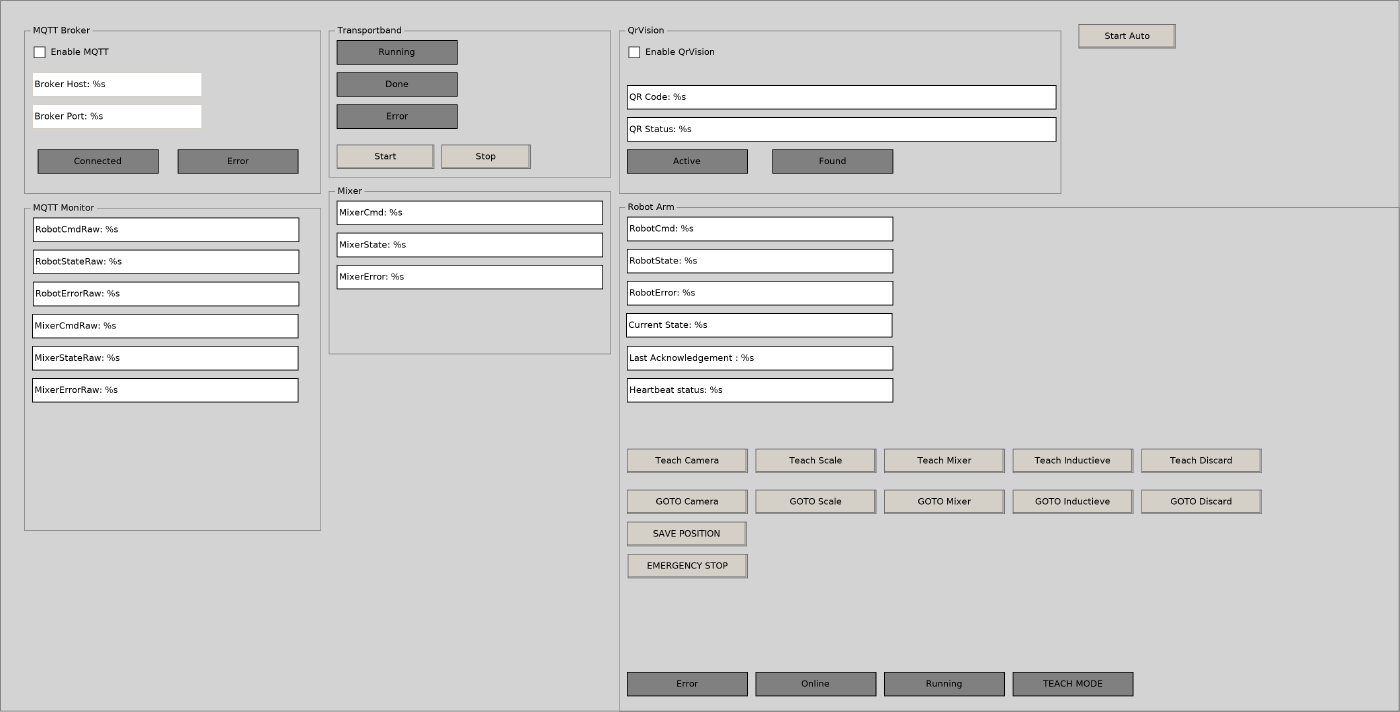
VISUALIZATION PannenkoekenDashboard  // 1742x887
    GroupBox (30,30 369x211), "MQTT Broker"
        Checkbox (10,20 150x30), "Enable MQTT", variable: GVL_MQTT.bEnableMqtt
        Rectangle (191,156 150x30), "Error"
        Rectangle (17,156 150x30), "Connected", colour toggle: GVL_MQTT.bMqttConnected
        Textfield (10,60 211x30), "Broker Host: %s", text variable: GVL_MQTT.sMqttBroker
        Textfield (10,100 211x30), "Broker Port: %s", text variable: GVL_MQTT.nMqttPort
    GroupBox (30,251 369x410), "MQTT Monitor"
        Rectangle (10,140 331x30), "MixerCmdRaw: %s", text variable: GVL_MQTT.sMixerCmdRaw
        Rectangle (10,180 331x30), "MixerStateRaw: %s", text variable: GVL_MQTT.sMixerStateRaw
        Rectangle (10,220 331x30), "MixerErrorRaw: %s", text variable: GVL_MQTT.sMixerErrorRaw
        Rectangle (11,20 331x30), "RobotCmdRaw: %s", text variable: GVL_MQTT.sRobotCmdRaw
        Rectangle (11,60 331x30), "RobotStateRaw: %s", text variable: GVL_MQTT.sRobotStateRaw
        Rectangle (11,100 331x30), "RobotErrorRaw: %s", text variable: GVL_MQTT.sRobotErrorRaw
    GroupBox (770,250 972x637), "Robot Arm"
        Rectangle (10,20 331x30), "RobotCmd: %s", text variable: GVL_MQTT.sRobotCmdDisplay
        Rectangle (10,60 331x30), "RobotState: %s", text variable: GVL_MQTT.sRobotStateDisplay
        Rectangle (10,100 331x30), "RobotError: %s", text variable: GVL_MQTT.sRobotErrorDisplay
        Rectangle (10,587 150x30), "Error", colour toggle: GVL_MQTT.bRobotArmAlarm
        Rectangle (170,587 150x30), "Online", colour toggle: GVL_MQTT.bRobotArmOnline
        Rectangle (330,587 150x30), "Running", colour toggle: GVL_MQTT.bRobotArmBusy
        Rectangle (10,221 331x30), "Heartbeat status: %s", text variable: GVL_MQTT.sRobotHeartbeatDisplay
        Rectangle (9,140 331x30), "Current State: %s", text variable: GVL_MQTT.sRobotArmDisplay
        Button (10,309 150x30), "Teach Camera"
            OnMouseClick: execute { GVL_MQTT.sRobotTargetPose := 'camera'; GVL_MQTT.bVisuRobotTeach  := TRUE; }
        Button (170,309 150x30), "Teach Scale"
            OnMouseClick: execute { GVL_MQTT.sRobotTargetPose := 'scale'; GVL_MQTT.bVisuRobotTeach  := TRUE; }
        Button (330,309 150x30), "Teach Mixer"
            OnMouseClick: execute { GVL_MQTT.sRobotTargetPose := 'mixer'; GVL_MQTT.bVisuRobotTeach  := TRUE; }
        Button (490,309 150x30), "Teach Inductieve"
            OnMouseClick: execute { GVL_MQTT.sRobotTargetPose := 'inductive'; GVL_MQTT.bVisuRobotTeach  := TRUE; }
        Button (650,309 150x30), "Teach Discard"
            OnMouseClick: execute { GVL_MQTT.sRobotTargetPose := 'discard'; GVL_MQTT.bVisuRobotTeach  := TRUE; }
        Button (10,360 150x30), "GOTO Camera"
            OnMouseClick: execute { GVL_MQTT.sRobotTargetPose := 'camera'; GVL_MQTT.bVisuRobotGoto   := TRUE; }
        Button (10,400 149x30), "SAVE POSITION"
            tap GVL_MQTT.bVisuRobotSave
        Button (11,440 149x30), "EMERGENCY STOP"
            tap GVL_MQTT.bVisuRobotStop
        Rectangle (10,181 331x30), "Last Acknowledgement : %s", text variable: GVL_MQTT.sRobotArmAck
        Rectangle (490,587 150x30), "TEACH MODE", colour toggle: GVL_MQTT.bRobotArmTeachMode
    GroupBox (409,30 351x191), "Transportband"
        Button (10,150 121x30), "Start"
            tap GVL_MQTT.bVisuStartTransportband
        Button (140,150 111x30), "Stop"
            tap GVL_MQTT.bVisuStopTransportband
        Rectangle (10,20 150x30), "Running", colour toggle: GVL_MQTT.bTransportbandRunning
        Rectangle (10,60 150x30), "Done", colour toggle: GVL_MQTT.bTransportbandDone
        Rectangle (10,100 150x30), "Error", colour toggle: GVL_MQTT.bSystemError
    GroupBox (409,230 351x211), "Mixer"
        Rectangle (10,60 331x30), "MixerState: %s", text variable: GVL_MQTT.sMixerStateDisplay
        Rectangle (10,20 331x30), "MixerCmd: %s", text variable: GVL_MQTT.sMixerCmdDisplay
        Rectangle (10,100 331x30), "MixerError: %s", text variable: GVL_MQTT.sMixerErrorDisplay
    GroupBox (770,30 550x211), "QrVision"
        Rectangle (10,76 534x30), "QR Code: %s", text variable: GVL_Data.sQrCodeText
        Rectangle (10,116 534x30), "QR Status: %s", text variable: GVL_Data.sQrDisplayText
        Rectangle (10,156 150x30), "Active", colour toggle: GVL_Data.bQrActive
        Rectangle (191,156 150x30), "Found", colour toggle: GVL_Data.bQrCodeFound
        Checkbox (10,20 150x30), "Enable QrVision", variable: GVL_Data.bQrEnabled
    Button (940,610 150x30), "GOTO Scale"
        OnMouseClick: execute { GVL_MQTT.sRobotTargetPose := 'scale'; GVL_MQTT.bVisuRobotGoto   := TRUE; }
    Button (1100,610 150x30), "GOTO Mixer"
        OnMouseClick: execute { GVL_MQTT.sRobotTargetPose := 'mixer'; GVL_MQTT.bVisuRobotGoto   := TRUE; }
    Button (1260,610 150x30), "GOTO Inductieve"
        OnMouseClick: execute { GVL_MQTT.sRobotTargetPose := 'inductive'; GVL_MQTT.bVisuRobotGoto   := TRUE; }
    Button (1420,610 150x30), "GOTO Discard"
        OnMouseClick: execute { GVL_MQTT.sRobotTargetPose := 'discard'; GVL_MQTT.bVisuRobotGoto   := TRUE; }
    Button (1342,30 121x30), "Start Auto"
        tap GVL_MQTT.bVisuStartSequence
END_VISUALIZATION

(* stored: Version 1.1.0.1, ProductVersion 3.1.4026.17
   Visu PannenkoekenDashboard: Id {747fc4aa-41f4-4f69-b086-b41493138125} *)
